{attribute 'qualified_only'}
VAR_GLOBAL CONSTANT
	// Program/logic safety limits
	DEFAULT_MAX_ATTRIBUTE_COUNT: 	UDINT := 20;  	// Maximum attributes for FB_Attributes
	DEFAULT_MAX_LINK_COUNT:			UDINT := 128;	// Maximum links a span keeps, the OpenTelemetry default
	MAX_LOOP_COUNT:					UDINT := 20000; // Maximum iterations a for/while loop can have
	MAX_LOG_RECORDS_PER_SCAN: 		UDINT := 100;  	// Maximum number of log records that can be emitted per scan.
	MAX_SPAN_RECORDS_PER_SCAN:		UDINT := 100;	// Maximum number of spans that can be emitted per scan.
END_VAR
VAR_GLOBAL
	_ID: UDINT := 1;
	defaultSampler: FB_Sampler;  // ParentBased(root=AlwaysOn); stateless, so providers share it
END_VAR

(* stored: Version 1.1.0.1
   GVL TcOtlp_GVL: Id {2c8a878d-5952-40c2-818b-cd6117aea204}
   Property NEXT_ID: Id {66a2dc14-5b7c-4295-87ce-3f72d7397f26}
   Get Get: Id {67ac250b-bd9e-4a04-b15e-fab6928fa6d3} *)
